GLOBALCONSTANTS logiBUS_ENC (* logiBUS_ENC constants *)
  (* Standard: 61499-1; Description: Copyright (c) 2026 HR Agrartechnik GmbH This program and the accompanying materials are made available under the terms of the Eclipse Public License 2.0 which is available at https://www.eclipse.org/legal/epl-2.0/ SPDX-License-Identifier: EPL-2.0 *)
  (* Version 1.0, 2026-11-26, Franz Höpfinger, HR Agrartechnik GmbH *)
  PACKAGE logiBUS::io::ENC;
  VAR_GLOBAL CONSTANT
    Encoder_E1 : logiBUS::io::ENC::logiBUS_ENC_S := (Pin := 1);
    Invalid : logiBUS::io::ENC::logiBUS_ENC_S := (Pin := 255);
  END_VAR
END_GLOBALCONSTANTS
